KUKA KRL program: Prog_Name_That_I.src

&ACCESS RVP
&REL 1
&PARAM TEMPLATE = C:\KRC\Roboter\Template\vorgabe
&PARAM EDITMASK = *
DEF Prog_Name_That_I ( )

; External program calls:
EXT Program_With_A_L()

EXT BAS (BAS_COMMAND :IN,REAL :IN )


; GLOBAL INTERRUPT DECL 3 WHEN $STOPMESS==TRUE DO IR_STOPM ( )
; INTERRUPT ON 3

;FOLD Initialise and set default speed
BAS (#INITMOV,0)
BAS (#VEL_PTP,100)
BAS (#ACC_PTP,20)
$VEL.CP=0.2
BAS (#TOOL,0)
BAS (#BASE,0)
;ENDFOLD

;;FOLD STARTPOS
;$BWDSTART = FALSE
;PDAT_ACT = PDEFAULT
;BAS(#PTP_DAT)
;FDAT_ACT = {TOOL_NO 0,BASE_NO 0,IPO_FRAME #BASE}
;BAS(#FRAMES)
;;ENDFOLD

$ADVANCE = 5

;FOLD ---- Quickly skip BCO ----
; PTP $AXIS_ACT
;ENDFOLD

;FOLD ---- GO HOME ----
; PTP {A1 0.000, A2 -90.000, A3 90.000, A4 0.000, A5 0.000, A6 0.000, E1 0, E2 0, E3 0, E4 0, E5 0, E6 0}
;ENDFOLD


; Program generated by VerticalBot Studio for KUKA KR 6 R900 sixx on 25/10/2026 12:00:00
; Using nominal kinematics.
; ---- Setting reference (Base) ----
$BASE = {FRAME: X 0.000,Y 0.000,Z 0.000,A 0.000,B 0.000,C 0.000}
; BASE_DATA[1] = {FRAME: X 0.000,Y 0.000,Z 0.000,A 0.000,B 0.000,C 0.000}
; $BASE = BASE_DATA[1]
; --------------------------
; ---- Setting tool (TCP) ----
$TOOL = {FRAME: X 10.000,Y 0.000,Z 120.000,A 0.000,B 15.000,C 0.000}
; --------------------------
$VEL.CP = 1.00000
$APO.CPTP = 10
$APO.CDIS = 10.000
PTP {A1 10.00000,A2 -80.00000,A3 100.00000,A4 20.00000,A5 40.00000,A6 -30.00000} C_PTP
LIN {X 549.094,Y 5.962,Z 504.960,A -174.431,B 15.001,C 175.695} C_DIS
$APO.CPTP = 0
$APO.CDIS = 0.500
LIN {X 506.272,Y -26.320,Z 503.226,A -178.509,B 14.048,C 175.384} C_DIS
HALT
WAIT SEC 1.500
Wait for StrClear($LOOP_MSG[])
$LOOP_CONT = TRUE
$LOOP_MSG[] = "Say "hi" to the operator"
; A long comment line that exceeds the usual controller limits for comments by far, really
$OUT[12]=FALSE
OUT_A=TRUE
START_TIMER:
$TIMER_STOP[1]=TRUE
$TIMER_FLAG[1]=FALSE
$TIMER[1]=1.000
$TIMER_STOP[1]=FALSE
WAIT FOR ($IN[4]==FALSE OR $TIMER_FLAG[1])
$TIMER_STOP[1]=TRUE
IF $TIMER_FLAG[1]== TRUE THEN
    HALT ; Timed out!
    GOTO START_TIMER
ENDIF
WAIT FOR (IN_B==TRUE)
Program_With_A_L()
; ---- Setting reference (Base) ----
; BASE_DATA[12] = {FRAME: X 250.000,Y 300.000,Z -10.000,A 90.000,B 0.000,C 0.000}
$BASE = {FRAME: X 250.000,Y 300.000,Z -10.000,A 90.000,B 0.000,C 0.000}
; $BASE = BASE_DATA[12]
; --------------------------
; ---- Setting tool (TCP) ----
; TOOL_DATA[7] = {FRAME: X 10.000,Y 0.000,Z 120.000,A 0.000,B 15.000,C 0.000}
$TOOL = {FRAME: X 10.000,Y 0.000,Z 120.000,A 0.000,B 15.000,C 0.000}
; $TOOL = TOOL_DATA[7]
; --------------------------
$VEL.ORI1 = 30.00000
$VEL.ORI2 = 30.00000
$ACC.ORI1 = 100.00000
$ACC.ORI2 = 100.00000
LIN {X 549.094,Y 5.962,Z 504.960,A -174.431,B 15.001,C 175.695} C_DIS
PTP {A1 10.00000,A2 -80.00000,A3 100.00000,A4 20.00000,A5 40.00000,A6 -30.00000}
END
